{region 'Documentation'}
(*!
<summary>Checks whether the INT value is outside the inclusive range.</summary>
<description>

Minimum &gt; Maximum reports Error during active evaluation; equal bounds are
valid.

</description>
*)
{endregion}
FUNCTION_BLOCK AssertNotInRange_Int EXTENDS AssertionBase
VAR_INPUT
    IN : INT; //! Actual value checked or observed by this Assertion.
    Minimum : INT; //! Inclusive lower bound of the comparison; for a range, must not exceed Maximum.
    Maximum : INT; //! Inclusive upper bound of the comparison; for a range, must not be below Minimum.
END_VAR

SUPER^();

{region 'Documentation'}
(*!
<summary>Check whether the INT value is outside the inclusive range.</summary>
*)
{endregion}
METHOD PROTECTED Assert
VAR
    Message : STRING(GVL_Constants.MessageLength);
    MinimumText : STRING(GVL_Constants.AssertionValueLength);
    MaximumText : STRING(GVL_Constants.AssertionValueLength);
    ActualText : STRING(GVL_Constants.AssertionValueLength);
END_VAR
IF NOT EvaluationActive THEN
    RETURN;
END_IF;

IF Result = E_Result.Error THEN
    RETURN;
END_IF;

IF Minimum > Maximum THEN
    MinimumText := INT_TO_STRING(Minimum);
    MaximumText := INT_TO_STRING(Maximum);
    Message := CONCAT('Assertion error: minimum exceeds maximum. Minimum = ',
        MinimumText);
    Message := CONCAT(Message, ', Maximum = ');
    Message := CONCAT(Message, MaximumText);
    Message := CONCAT(Message, '.');
    Error(Message := Message);
    RETURN;
END_IF;

IF Result = E_Result.Failed THEN
    RETURN;
END_IF;

IF (IN >= Minimum) AND (IN <= Maximum) THEN
    MinimumText := INT_TO_STRING(Minimum);
    MaximumText := INT_TO_STRING(Maximum);
    ActualText := INT_TO_STRING(IN);
    Message := CONCAT('Assertion failed: value is inside forbidden range. Minimum = ',
        MinimumText);
    Message := CONCAT(Message, ', Maximum = ');
    Message := CONCAT(Message, MaximumText);
    Message := CONCAT(Message, ', Actual = ');
    Message := CONCAT(Message, ActualText);
    Message := CONCAT(Message, '.');
    Fail(Message := Message);
    RETURN;
END_IF;

Pass();
END_METHOD

END_FUNCTION_BLOCK

(* stored: Version 1.1.0.1
   POU AssertNotInRange_Int: Id {0f20f7d3-d159-4478-bd93-78484475cf76}, SpecialFunc None
   Folder Internal: Id {1e6bbc67-54cb-4c4e-ac49-b1ef7ec5ffae}
   Method Assert: Id {de3e1ab4-ea69-46e7-9b19-b0acdd275738} *)
